(* IEC 61131-3 sources: Elmo_Master/Lasal_PRG/Welcon8Axis_EtherCAT_Test_With_RobotAxis/Class/EtherCAT_Hub_Base, 1 file *)

(* ---- EtherCAT_Hub_Base.st ---- *)
#include "..\..\Class\ECAT_Master_Base\ECAT_Master_Base.h"
#include "..\..\Source\interfaces\lsl_st_hardwaretree.h"

(*!
<Class
	Name               = "EtherCAT_Hub_Base"
	Revision           = "1.2"
	RealtimeTask       = "false"
	CyclicTask         = "false"
	BackgroundTask     = "false"
	Sigmatek           = "true"
	OSInterface        = "false"
	HighPriority       = "false"
	Automatic          = "false"
	UpdateMode         = "Prescan"
	IconPath           = ".\Class\EtherCAT.ico"
	SharedCommandTable = "true"
	Objectsize         = "(494,120)">
	<Channels>
		<Server Name="ClassSvr" Visualized="false" Initialize="false" WriteProtected="true" Retentive="false" Comment="Connect an EtherCAT Slave."/>
		<Client Name="BusType" Required="false" Internal="false" DefValue="0" Comment="Type of the Bus&#13;&#10;0 .. EtherCAT&#13;&#10;1 .. LVDS&#13;&#10;Else .. Not supported&#13;&#10;"/>
		<Client Name="SplitterPlace" Required="true" Internal="false" Comment="Place of this splitter."/>
		<Client Name="toNextEtherCAT" Required="true" Internal="false" Comment="Connect to first server of Ethercat master."/>
	</Channels>
	<Dependencies>
		<Files>
			<File Path=".\Class\ECAT_Master_Base\ECAT_Master_Base.h" Include="true"/>
			<File Path=".\Source\interfaces\lsl_st_hardwaretree.h" Include="true"/>
		</Files>
	</Dependencies>
	<RevDoku>
		<Owner Company="Sigmatek" Author="EisMic"/>
		<Dokumentation Revision="1.2" Date="2026-04-10" Author="LanSte" Company="Sigmatek" Description="Special: Set property flag &quot;Hidden&quot; of class, since this is an internal class."/>
		<Dokumentation Revision="1.1" Date="27.05.2024" Author="LanSte" Company="Sigmatek" Description="Added Support for HW-Paths and LVDS Bus."/>
		<Dokumentation Revision="1.0" Date="09.04.2020" Author="EisMic" Company="Sigmatek" Description="First release version"/>
		<Dokumentation Revision="0.1" Date="17.05.2019" Author="EisMic" Company="Sigmatek" Description="First test version."/>
	</RevDoku>
	<AdditionalData>
		<Entry Name="Hidden" Value="true"/>
	</AdditionalData>
</Class>
*)
EtherCAT_Hub_Base : CLASS
  //Servers:
	ClassSvr 	: SvrChCmd_DINT;
  //Clients:
	toNextEtherCAT 	: CltChCmd_t_e_VaranErrors;
	SplitterPlace 	: CltCh_DINT;
	BusType 	: CltCh_DINT;
  //Variables:
  //Functions:

	FUNCTION VIRTUAL GLOBAL ClassSvr::NewInst
		VAR_INPUT
			pPara 	: ^CmdStruct;
			pResult 	: ^results;
		END_VAR
		VAR_OUTPUT
			ret_code 	: iprStates;
		END_VAR;
  //Tables:
	FUNCTION @STD
		VAR_OUTPUT
			ret_code	: CONFSTATES;
		END_VAR;
	FUNCTION GLOBAL TAB @CT_;
END_CLASS;

FUNCTION VIRTUAL GLOBAL EtherCAT_Hub_Base::ClassSvr::NewInst
	VAR_INPUT
		pPara 	: ^CmdStruct;
		pResult 	: ^results;
	END_VAR
	VAR_OUTPUT
		ret_code 	: iprStates;
	END_VAR

  case pPara^.uiCmd of

//**********************************************************************************************************************************************************
    ECAT_M_GET_HW_PATH:

      ret_code := toNextEtherCAT.NewInst(pPara, pResult);
      if (ret_code = READY) & (pResult^.aData[4]$DINT = 2) then // Result Ok and Version = 2

        // Insert Escape Sequence into result
        if BusType = 0 then
          pResult^.aData[12]$HSINT  := HWT_ESCAPE_ECAT;
        elsif BusType = 1 then
          pResult^.aData[12]$HSINT  := HWT_ESCAPE_ECAT_LVDS;
        else
          ret_code := ERROR;
          pResult^.aData[0]$DINT    := ECAT_RETERR_CMD_INVALID_HWPATH_ESCAPE_SEQU;
          pResult^.aData[12]$HSINT  := HWT_ESCAPE_SEQU; // Unkown!
        end_if;

        pResult^.aData[13]$USINT  := SplitterPlace$USINT;

      end_if;

  else
    ret_code := toNextEtherCAT.NewInst(pPara, pResult);
  end_case;

END_FUNCTION
